        | 	local end_rel = pose_trans(pose_inv(p_center), scoop_end_pose)
        | 	local end_rel_tilted = pose_trans(end_rel, p[0, 0, 0, 0, ry, 0])
        | 	global tilted_pose_in_base = pose_trans(p_center, p[0,correction_y,correction_z,end_rel_tilted[3],end_rel_tilted[4], end_rel_tilted[5]])
        | 	global tilted_pose_in_base = pose_trans(tilted_pose_in_base, p[0, 0, spatula_len, 0, 0, 0])
        | 
        | 	if (Pow_name == "lactose_fine" or Pow_name == "Magnesium_sterate"):
        | 		tilt_send((angle_deg+5))
        | 	end
        | 	movel(tilted_pose_in_base, a=0.03, v=0.1)
        | 
        | 	if (Pow_name == "lactose_fine" or Pow_name == "Magnesium_sterate"):
        | 		tilt_send((angle_deg-5))
        | 	end
        | 
        | 	if (spatula=="spatula_flat_S" or spatula=="spatula_S"):
        | 		vibration_3()
        | 	else:
        | 		set_analog_out(0, vibration_voltage)
        | 	end
        | 	if (Pow_name=="Mannitol" or Pow_name =="NaCl"):
        | 		local n=1.4
        | 	else:
        | 		local n=1.5
        | 	end
        | 	local ry_level = deg2rad(ry_deg/n)
        | 	local end_rel_tilted_level = pose_trans(end_rel, p[0, 0, 0, 0, ry_level, 0])
        | 	local level_tilted_pose_in_base = pose_trans(p_center, p[0,correction_y,correction_z,end_rel_tilted_level[3],end_rel_tilted_level[4], end_rel_tilted_level[5]])
        | 	local level_tilted_pose_in_base = pose_trans(level_tilted_pose_in_base, p[0, 0, spatula_len, 0, 0, 0])
        | 
        | 	movel(level_tilted_pose_in_base, a=0.03, v=0.1)
        | 	#if (level>70.0):
        | 		#sleep(1.0)
        | 	#end
        | 	sleep(1.0)
        | 	#sleep(vibration_time)
        | 
        | 	movel(tilted_pose_in_base, a=0.03, v=0.1)
        | 	set_analog_out(0, 0.0)
        | 
        | 	tilt_pose_rel = pose_trans(pose_inv(p_center), tilted_pose_in_base)
        | 
        | 	lifted_pose_rel = pose_trans(lift_offset, tilt_pose_rel)
        | 
        | 	global lifted_pose = pose_trans(p_center, lifted_pose_rel)
        | 	movel(lifted_pose, a=0.03, v=0.1)
        | 	CCW_Rotate()
        | end
        | 
        | 
        | # calculate center pose on top of the container using pose transformation
        | def center_pose():
        | 	# pose transformation from side of the container to top to get center point
        | 	trans_rel = p[-0.005, 0.05, -0.027, 0, 0, 0]
        | 
        | 	p_translated = pose_trans(place_pose, trans_rel)
        | 	cx = p_translated[0]
        | 	cy = p_translated[1]
        | 	cz = p_translated[2]
        | 
        | 	global p_center_vertical = p[cx,cy,cz, 0, 0, 4.14]
        | 
        | 	#movej(p_center_vertical, a =0.3, v =0.3)
        | 	return p_center_vertical
        | end
        | 
        | # update center pose based on tilting
        | def updated_center_pose(p_center_vertical, angle_deg):
        | 	hinge_pose = pose_trans(p_center_vertical, p[0,0,-0.2,0,0,0])
        | 	local_rel = pose_trans(pose_inv(hinge_pose), p_center_vertical)
        | 
        | 	rot_tilt = p[0,0,0, -deg2rad(angle_deg),0,0]
        | 	local_rel_tilted = pose_trans(rot_tilt, local_rel)
        | 
        | 	global p_center = pose_trans(hinge_pose, local_rel_tilted)
        | 	return p_center
        | end
        | 
        | #------
        | # POTS commands
        | def tilt_send(angle):
        | 	socket_open("192.168.12.101", 80)
        | 	angle = 92.0 - angle
        | 	socket_send_string("Tilt,"+to_str(angle)+",0")
        | 	sync()
        | 	sleep(0.5)
        | 	socket_close()
        | end
        | 
        | def Motors_off():
        | 	socket_open("192.168.12.101", 80)
        | 	socket_send_string("Off,0,0")
        | 	sync()
        | 	sleep(0.5)
        | 	socket_close()
        | end
        | 
        | def Rotate():
        | 	socket_open("192.168.12.101", 80)
        | 	socket_send_string("FullRotation, 1, 2000")
        | 	sync()
        | 	sleep(0.5)
        | 	socket_close()
        | end
        | 
        | 
        | def CCW_Rotate():
        | 	socket_open("192.168.12.101", 80)
        | 	socket_send_string("FullRotation, -1, 2000")
        | 	sync()
        | 	sleep(0.5)
        | 	socket_close()
        | end
        | 
        | def tilt_to_home():
        | 	socket_open("192.168.12.101", 80)
        | 	socket_send_string("Home,0,0")
        | 	sync()
        | 	sleep(0.5)
        | 	socket_close()
        | end
    SuppressedNode
      Script file /programs/04 Scripts/dosing.script
        | def vibration_2():
        | 	set_analog_out(0,0.4)
        | 	sleep(0.8)
        | 	set_analog_out(0,0.0)
        | 	sleep(0.2)
        | end
        | 
        | def vibration_3():
        | 	set_analog_out(0,0.4)
        | 	sleep(0.5)
        | 	set_analog_out(0,0.0)
        | 	sleep(0.3)
        | end
        | 
        | def vibration_4():
        | 	set_analog_out(0,0.4)
        | 	sleep(0.6)
        | 	set_analog_out(0, 0.0)
        | 	sleep(0.5)
        | end
        | 
        | def vibration_1():
        | 	set_analog_out(0,0.4)
        | 	sleep(1)
        | 	set_analog_out(0,0.0)
        | 	sleep(0)
        | end
        | 
        | def move_tilt_in_steps(Pow_center, final_pose, steps):
        | 	i = 0
        | 	while i <= steps:
        | 		ratio = i / steps
        | 		pose_step = p[Pow_center[0] + ratio * (final_pose[0] - Pow_center[0]), Pow_center[1] + ratio * (final_pose[1] -Pow_center[1]),Pow_center[2] + ratio * (final_pose[2] - Pow_center[2]), Pow_center[3] + ratio * (final_pose[3] - Pow_center[3]), Pow_center[4] + ratio * (final_pose[4] - Pow_center[4]), Pow_center[5] + ratio * (final_pose[5] - Pow_center[5])]
        | 		movej(pose_step, a=1.2, v=0.15)
        | 		sleep(0.1)
        | 		i = i+1
        | 	end
        | end
        | 
        | def tilt_container(angle):
        | 	p_center = get_actual_tcp_pose()
        | 	hinge_offset = p[0,0,-0.23,0,0,0]
        | 	pivot_pose = pose_trans(p_center, hinge_offset)
        | 	pose_rel = pose_trans(pose_inv(pivot_pose), p_center)
        | 	angle_mid = (angle/2.0)*3.1416/180
        | 	angle_end = angle*3.1416/180
        | 	tilt_mid = p[0,0,0, -angle_mid, 0, 0]
        | 	tilt_end = p[0,0,0, -angle_end, 0, 0]
        | 	pose_rel_mid = pose_trans(tilt_mid, pose_rel)
        | 	pose_rel_end = pose_trans(tilt_end, pose_rel)
        | 	via_pose = pose_trans(pivot_pose, pose_rel_mid)
        | 	end_pose = pose_trans(pivot_pose, pose_rel_end)
        | 	movec(via_pose, end_pose, a=0.05, v=0.01, r=0.001)
        | 	p_center = get_actual_tcp_pose()
        | end
        | 
        | def deg2rad(d):
        | 	return d*3.141592/180
        | end
        | 
        | def map_tilt_to_ry_deg(container_deg):
        | 	#ry_deg = -0.875*container_deg +87.0
        | 	#return clamp(ry_deg, 5.0, 80.0)
        | 	if (Pow_name == "NaCl" or Pow_name == "Mannitol" or Pow_name == "CCS" or Pow_name == "MCC"):
        | 		if ( level>=10.0):
        | 			ry_min = 10.0
        | 			ry_max = 75.0
        | 		elif (level<10.00 and level >1.00):
        | 			ry_min = 16.0
        | 			ry_max = 65.0
        | 		else:
        | 			ry_min=17.0
        | 			ry_max=75.0
        | 		end
        | 	else:
        | 		if ( level>=10.0):
        | 			ry_min = 0.0
        | 			ry_max = 65.0
        | 		elif (level<10.00 and level >1.00):
        | 			ry_min = 10.0
        | 			ry_max = 45.0
        | 		else:
        | 			ry_min=0.0
        | 			ry_max=50.0
        | 		end
        | 
        | 	end
        | 	local span_count = angle_max -angle_min
        | 	local span_ry = ry_max - ry_min
        | 
        | 	local t = (container_deg -angle_min)/span_count
        | 	local ry_deg = ry_max - t*span_ry
        | 
        | 	return clamp(ry_deg, ry_min, ry_max)
        | 
        | end
        | 
        | def caluclate_corrections(level):
        | 	z_high = 0.01
        | 	z_low = -0.08
        | 	y_high = -0.01
        | 	y_low = -0.015
        | 
        | 	scale = (level - 10.0) / (100.0-10.0)
        | 
        | 	global correction_z = z_low + scale*(z_high - z_low)
        | 	global correction_y = y_low + scale*(y_high -y_low)
        | 
        | end
        | 
        | def scoop_powder(p_center):
        | 	#lift_offset = p[0, 0, 0.05, 0, 0, 0]
        | 	vibration_voltage = 0.4
        | 	vibration_time = 3.0
        | 	diameter = 0.07
        | 	global scoop_radius_default = 0.0
        | 	#p_center = center_pose_t
        | 
        | 
        | 	if (level >=70.00):
        | 		approach_offset = p[0.008,0,0.22,0,0,0]
        | 		lift_offset = p[0, 0, 0.05, 0, 0, 0]
        | 		caluclate_corrections(level)
        | 	elif (level >=10.00 and level <70):
        | 		approach_offset = p[0.008,0,0.22,0,0,0]
        | 		lift_offset = p[0, 0, 0.15, 0, 0, 0]
        | 		caluclate_corrections(level)
        | 	elif (level<10.00 and level >= 1.00):
        | 		approach_offset = p[0.01,0,0.22,0,0,0]
        | 		correction_z = -0.08
        | 		correction_y = -0.01
        | 		lift_offset = p[0, 0, 0.14, 0, 0, 0]
        | 	else:
        | 		approach_offset = p[0.008,0,0.22,0,0,0]
        | 		correction_z = -0.08
        | 		correction_y = -0.01
        | 		lift_offset = p[0, 0, 0.14, 0, 0, 0]
        |  	end
        | 
        | 	if (spatula == "spatula_L"):
        | 		global spatula_depth = 0.015
        | 	elif (spatula == "spatula_M"):
        | 		global spatula_depth = 0.01
        | 	elif (spatula == "spatula_S"):
        | 		global spatula_depth = 0.008
        | 	elif (spatula == "spatula_flat_M"):
        | 		global spatula_depth = 0.001
        | 	elif (spatula == "spatula_flat_S"):
        | 		global spatula_depth = 0.005
        | 	end
        | 
        | 	scoop_radius_default = diameter/2 - spatula_depth
        | 	scoop_entry_pose = pose_trans(p_center, approach_offset)
        | 	movel(scoop_entry_pose, a=0.1, v=0.25)
        | 
        | 	scoop_start_rel = p[scoop_radius_default, 0, scoop_depth, 0, 0, 0]
        | 
        | 	rot_mid = p[0, 0, 0, 0, 0, 0.785]
        | 	rot_end = p[0, 0, 0, 0, 0, 1.5708]
        | 
        | 	scoop_via_rel = pose_trans(rot_mid, scoop_start_rel)
        | 	scoop_end_rel = pose_trans(rot_end, scoop_start_rel)
        | 
        | 	scoop_start_pose = pose_trans(p_center, scoop_start_rel)
        | 	scoop_via_pose = pose_trans(p_center, scoop_via_rel)
        | 	scoop_end_pose = pose_trans(p_center, scoop_end_rel)
        | 
        | 	movel(scoop_start_pose, a=0.5, v=0.3)
        | 	#movel(p_center, a=0.5, v=1.0)
        | 	#sleep(5.0)
        | 
        | 	if (level<90.0):
        | 		Rotate()
        | 	end
        | 
        | 	#movec(scoop_via_pose, scoop_end_pose, a=0.03, v=0.05)
        | 	movec(scoop_via_pose, scoop_end_pose, a=0.03, v=0.02)
        | 	#movel(pose_trans(get_actual_tcp_pose(), p[0,0,0,0,0,deg2rad(90.0)]), a=0.03, v=0.05)
        | 	sleep(1.0)
        | 	local ry_deg = map_tilt_to_ry_deg(angle_deg)
        | 	local ry = deg2rad(ry_deg)
        | 	local end_rel = pose_trans(pose_inv(p_center), scoop_end_pose)
        | 	local end_rel_tilted = pose_trans(end_rel, p[0, 0, 0, 0, ry, 0])
        | 	global tilted_pose_in_base = pose_trans(p_center, p[0,correction_y,correction_z,end_rel_tilted[3],end_rel_tilted[4], end_rel_tilted[5]])
        | 	global tilted_pose_in_base = pose_trans(tilted_pose_in_base, p[0, 0, spatula_len, 0, 0, 0])
        | 
        | 	if (Pow_name == "lactose_fine" or Pow_name == "Magnesium_sterate"):
        | 		tilt_send((angle_deg+5))
        | 	end
        | 	movel(tilted_pose_in_base, a=0.03, v=0.1)
        | 
        | 	if (Pow_name == "lactose_fine" or Pow_name == "Magnesium_sterate"):
        | 		tilt_send((angle_deg-5))
        | 	end
        | 
        | 	if (spatula=="spatula_flat_S" or spatula=="spatula_S"):
        | 		vibration_3()
        | 	else:
        | 		set_analog_out(0, vibration_voltage)
        | 	end
        | 	if (Pow_name=="Mannitol" or Pow_name =="NaCl"):
        | 		local n=1.4
        | 	else:
        | 		local n=1.5
        | 	end
        | 	local ry_level = deg2rad(ry_deg/n)
        | 	local end_rel_tilted_level = pose_trans(end_rel, p[0, 0, 0, 0, ry_level, 0])
        | 	local level_tilted_pose_in_base = pose_trans(p_center, p[0,correction_y,correction_z,end_rel_tilted_level[3],end_rel_tilted_level[4], end_rel_tilted_level[5]])
        | 	local level_tilted_pose_in_base = pose_trans(level_tilted_pose_in_base, p[0, 0, spatula_len, 0, 0, 0])
        | 
        | 	movel(level_tilted_pose_in_base, a=0.03, v=0.1)
        | 	#if (level>70.0):
        | 		#sleep(1.0)
        | 	#end
        | 	sleep(1.0)
        | 	#sleep(vibration_time)
        | 
        | 	movel(tilted_pose_in_base, a=0.03, v=0.1)
        | 	set_analog_out(0, 0.0)
        | 
        | 	tilt_pose_rel = pose_trans(pose_inv(p_center), tilted_pose_in_base)
        | 
        | 	lifted_pose_rel = pose_trans(lift_offset, tilt_pose_rel)
        | 
        | 	global lifted_pose = pose_trans(p_center, lifted_pose_rel)
        | 	movel(lifted_pose, a=0.03, v=0.1)
        | 	CCW_Rotate()
        | end
        | 
        | 
        | def center_pose():
        | 	trans_rel = p[-0.005, 0.05, -0.015, 0, 0, 0]
        | 
        | 	p_translated = pose_trans(place_pose, trans_rel)
        | 	cx = p_translated[0]
        | 	cy = p_translated[1]
        | 	cz = p_translated[2]
        | 
        | 	global p_center_vertical = p[cx,cy,cz, 0, 0, 4.09]
        | 
        | 	#movej(p_center_vertical, a =0.3, v =0.3)
        | 	return p_center_vertical
        | end
        | 
        | def updated_center_pose(p_center_vertical, angle_deg):
        | 	hinge_pose = pose_trans(p_center_vertical, p[0,0,-0.2,0,0,0])
        | 	local_rel = pose_trans(pose_inv(hinge_pose), p_center_vertical)
        | 
        | 	rot_tilt = p[0,0,0, -deg2rad(angle_deg),0,0]
        | 	local_rel_tilted = pose_trans(rot_tilt, local_rel)
        | 
        | 	global p_center = pose_trans(hinge_pose, local_rel_tilted)
        | 	return p_center
        | end
        | 
        | def tilt_send(angle):
        | 	socket_open("192.168.12.101", 80)
        | 	angle = 92.0 - angle
        | 	socket_send_string("Tilt,"+to_str(angle)+",0")
        | 	sync()
        | 	sleep(0.5)
        | 	socket_close()
        | end
        | 
        | def Motors_off():
        | 	socket_open("192.168.12.101", 80)
        | 	socket_send_string("Off,0,0")
        | 	sync()
        | 	sleep(0.5)
        | 	socket_close()
        | end
        | 
        | def Rotate():
        | 	socket_open("192.168.12.101", 80)
        | 	socket_send_string("FullRotation, 1, 2000")
        | 	sync()
        | 	sleep(0.5)
        | 	socket_close()
        | end
        | 
        | 
        | def CCW_Rotate():
        | 	socket_open("192.168.12.101", 80)
        | 	socket_send_string("FullRotation, -1, 2000")
        | 	sync()
        | 	sleep(0.5)
        | 	socket_close()
        | end
        | def tilt_to_home():
        | 	socket_open("192.168.12.101", 80)
        | 	socket_send_string("Home,0,0")
        | 	sync()
        | 	sleep(0.5)
        | 	socket_close()
        | end
    Script file /programs/04 Scripts/Powder_all.script
      | global SERVER_IP   = "192.168.12.139"
      | global SERVER_PORT = 3002
      | 
      | global container_id = 0
      | global powder_id  = 0
      | global bulk_density = 0
      | global H          = 0
      | global H_c          = 0
      | global mouth_d     = 0
      | global mouth_sh    = 0
      | global length_c     = 0
      | global diameter   = 0
      | global empty_weight_g  = 0
      | global volume_ml    = 0
      | global shape_code   = 0
      | global flow_code   = 0
      | global shape = ""
      | global Flowability = ""
      | global full_weight_g = 0
      | global cent_edge = 0
      | global pick_2_base = 0.2 # distance from tcp to base of picking table
      | global wall_thickness = 0.001
      | 
      | def read_db_data():
      | 
      |   socket_open(SERVER_IP, SERVER_PORT)
      |   sleep(0.5)
      |   socket_send_string("GET_DATACODE_FLOATS")
      |   sleep(5)
      | 
      |   local fl = socket_read_ascii_float(14)
      |   socket_close()
      | 
      |   global container_id = fl[1]
      |   global powder_id = fl[2]
      |   global bulk_density = fl[3]
      |   global H          = fl[4]/1000
      |   global H_c          = fl[5]/1000
      |   global mouth_d     = fl[6]/1000
      |   global mouth_sh    = fl[7]/1000
      |   global length_c     = fl[8]/1000
      |   global diameter   = fl[9]/1000
      |   global empty_weight_g = fl[10]
      |   global volume_ml    = fl[11]
      |   global full_weight_g = fl[12]
      |   global flow_code   = fl[13]
      |   global shape_code   = fl[14]
      | 
      | 	if (flow_code == 1.0):
      | 	  global Flowability = "MEDIUM"
      | 	elif (flow_code == 2.0):
      | 	  global Flowability = "LOW"
      | 	else:
      | 	  global Flowability = "HIGH"
      | 	end
      | 
      |   if ( shape_code == 1.0):
      | 	shape = "cylindrical"
      | 	cent_edge =  diameter
      |   else:
      | 	shape = "cubical"
      | 	cent_edge =  length_c
      |   end
      | 
      | end
      | 
      | 
      | def send_picking_info(Pow_name, target_weight):
      |   socket_open(SERVER_IP, SERVER_PORT)
      |   cmd = "PICK:"+Pow_name+";"+to_str(target_weight)
      |   socket_send_string(cmd)
      |   sleep(0.1)
      |   socket_close()
      | end
      | 
      | #### POTS ####
      | def tilt_send(angle):
      | 	socket_open("192.168.12.101", 80)
      | 	angle = 90.0 - angle
      | 	socket_send_string("Tilt,"+to_str(angle)+",0")
      | 	sync()
      | 	sleep(0.5)
      | 	socket_close()
      | end
      | 
      | def Motors_off():
      | 	socket_open("192.168.12.101", 80)
      | 	socket_send_string("Off,0,0")
      | 	sync()
      | 	sleep(0.5)
      | 	socket_close()
      | end
      | 
      | def Rotate():
      | 	socket_open("192.168.12.101", 80)
      | 	socket_send_string("FullRotation, 1, 2000")
      | 	sync()
      | 	sleep(0.5)
      | 	socket_close()
      | end
      | 
      | def CCW_Rotate():
      | 	socket_open("192.168.12.101", 80)
      | 	socket_send_string("FullRotation, -1, 2000")
      | 	sync()
      | 	sleep(0.5)
      | 	socket_close()
      | end
      | 
      | def tilt_to_home():
      | 	socket_open("192.168.12.101", 80)
      | 	socket_send_string("Home,0,0")
      | 	sync()
      | 	sleep(0.5)
      | 	socket_close()
      | end
      | #######
      | def vibration_1():
      | 	set_analog_out(0,0.4)
      | 	sleep(1)
      | 	set_analog_out(0,0.0)
      | 	sleep(0)
      | end
      | 
      | def vibration_2():
      | 	set_analog_out(0,0.4)
      | 	sleep(0.8)
      | 	set_analog_out(0,0.0)
      | 	sleep(0.2)
      | end
      | 
      | def vibration_3():
      | 	set_analog_out(0,0.4)
      | 	sleep(0.5)
      | 	set_analog_out(0,0.0)
      | 	sleep(0.3)
      | end
      | 
      | def vibration_4():
      | 	set_analog_out(0,0.8)
      | 	sleep(0.6)
      | 	set_analog_out(0, 0.0)
      | 	sleep(0.5)
      | end
      | 
      | ##################
      | 
      | global gear_2_holder = 0.018
      | global gain_per_percent = 0.5
      | global w_dosed_total = 0.0
      | global last_scale = 0.0
      | global tilt_angle_sent = 0.0
      | global level = 0.0
      | global target_g = 0.0
      | global angle_max = 60
      | global angle_min = 10
      | global hinge_2_base = 0.0421
      | global TCP_2_tip_x = 0.0047
      | global spatula_len = 0.182
      | global spatula_offset = p[TCP_2_tip_x,0,spatula_len,0,0,0]
      | global SPATULA_L_VOL_ML = 5.0        # 1 teaspoon = 5 mL
      | global SPATULA_M_VOL_ML = 1.25       # 1/4 teaspoon = 1.25 mL
      | global SPATULA_S_VOL_ML = 0.15625    # 1/32 teaspoon = 0.15625 mL
      | global SPATULA_FLAT_M_VOL_ML  = 2.2
      | global SPATULA_FLAT_S_VOL_ML  = 1.2   #based on caluclations using rho = m/V
      | global ry_deg_safe = 0
      | global ry_deg = 0
      | 
      | 
      | 
      | def clamp(x, lo, hi):
      | 	if(x<lo):
      | 		return lo
      | 	elif (x>hi):
      | 		return hi
      | 	else:
      | 		return x
      | 	end
      | end
      | 
      | def compute_level_percent(W_now, weight_value):   # W_now = container+powder, weight_value = live scale reading
      |     local delta = weight_value - last_scale
      | 
      |     if (delta < 0.0):
      |         delta = 0.0
      |     end
      | 
      |     global w_dosed_total = w_dosed_total + delta
      |     global last_scale = weight_value     # update the last scale reading
      | 
      |     local W_eff = W_now - w_dosed_total
      |     if (W_eff <  empty_weight_g):
      |         W_eff =  empty_weight_g
      |     end
      | 
      |     # Compute powder level %
      |     level = 100.0 * (W_eff -  empty_weight_g) / (full_weight_g -  empty_weight_g)
      | 
      |     # Clamp to 0–100
      |     level = clamp(level, 0, 100)
      |   textmsg("deb 1 = ", level)
      |     return level
      | end
      | 
      | def deg2rad(d):
      | 	return d*3.141592/180
      | end
      | 
      | def my_abs(val):
      | 	if (val<0):
      | 		return -val
      | 	else:
      | 		return val
      | 	end
      | end
      | 
      | def compute_tilt_deg(level_percent):
      | 	angle = angle_min + gain_per_percent*(100.0-level_percent)
      | 
      |   	textmsg("deb 2 = ", angle)
      | 	return clamp(angle, angle_min, angle_max)
      | end
      | 
      | def tilt(level_percentage):
      | 	new_angle = compute_tilt_deg(level_percentage)
      | 	global angle_rel = new_angle - tilt_angle_sent
      | 
      | 	if my_abs(angle_rel)>2.0:
      | 		tilt_send(new_angle)
      | 		global angle_deg = new_angle
      | 		global tilt_angle_sent = new_angle
      | 		global p_center_vertical = center_pose()
      | 		global p_center = updated_center_pose(p_center_vertical, angle_deg)
      | 	end
      | 
      | 	if (level_percentage<85.0):
      | 		tilt_send(angle_deg)
      | 	end
      | end
      | 
      | def compute_scoop_depth(level):
      |   return ((100.0-level)/100.0)*(H -mouth_sh )
      | end
      | 
      | def map_tilt_to_ry_deg(container_deg, level):
      | 
      | 	if (Flowability == "HIGH" or Flowability == "MEDIUM"):
      | 		global scoop_depth = compute_scoop_depth(level)
      | 		safe_scoop_pivot = (mouth_d  - spatula_depth)/(scoop_depth+mouth_sh )
      | 		global ry_deg_safe = asin(safe_scoop_pivot)
      | 		global ry_deg = 90-container_deg
      | 	else:
      | 		global scoop_depth = compute_scoop_depth(level)
      | 		safe_scoop_pivot = (mouth_d  - spatula_depth)/(scoop_depth+mouth_sh )
      | 		global ry_deg_safe = asin(safe_scoop_pivot)
      | 		global ry_deg = 90-container_deg
      | 	end
      | 	return [ry_deg_safe,ry_deg]
      | end
      | 
      | def get_scoop_weight(spatula, bulk_density):
      | 
      | 	local vol = 0
      | 
      | 	if (spatula == "spatula_L"):
      | 		vol = SPATULA_L_VOL_ML
      | 		global spatula_depth = 0.015
      | 		global spatula_mid   = 0.016
      | 		global spatula_ry    = 0.0
      | 
      | 	elif (spatula == "spatula_M"):
      | 		vol = SPATULA_M_VOL_ML
      | 		global spatula_depth = 0.010
      | 		global spatula_mid   = 0.0105
      | 		global spatula_ry    = 0.0
      | 
      | 	elif (spatula == "spatula_S"):
      | 		vol = SPATULA_S_VOL_ML
      | 		global spatula_depth = 0.008
      | 		global spatula_mid   = 0.0063
      | 		global spatula_ry    = 0.0
      | 
      | 	elif (spatula == "spatula_flat_M"):
      | 		vol = SPATULA_FLAT_M_VOL_ML
      | 		global spatula_depth = 0.001
      | 		global spatula_mid   = 0.002
      | 		global spatula_ry    = 10.0
      | 
      | 	elif (spatula == "spatula_flat_S"):
      | 		vol = SPATULA_FLAT_S_VOL_ML
      | 		global spatula_depth = 0.005
      | 		global spatula_mid   = 0.016
      | 		global spatula_ry    = 2.0
      | 
      | 	else:
      | 		textmsg("Unknown spatula type")
      | 		return 0.0
      | 	end
      | 	global target_g = vol * bulk_density
      | 	return target_g
      | 
      | end
      | 
      | def select_spatula(Flowability, level, diff, bulk_density, mouth_d ):
      | 
      |     local k = 1.1
      | 
      |     global powder_height = (H  - mouth_sh ) * level/100
      | 
      |     # =====================================================
      |     # LOW FLOWABILITY
      |     # =====================================================
      |     if (Flowability == "LOW"):
      | 
      |         local gFM = get_scoop_weight("spatula_flat_M", bulk_density)
      | 
      |         local level_ok_FM = (spatula_mid * 2 < powder_height)
      |         local diff_ok_FM  = (diff > k * gFM)
      | 
      |         local flatM_ok = level_ok_FM and diff_ok_FM
      | 
      |         if (flatM_ok):
      |             return "spatula_flat_M"
      |         else:
      |             return "spatula_flat_S"
      |         end
      | 
      |     end
      | 
      | 
      |     # =====================================================
      |     # LARGE
      |     # =====================================================
      |     local gL = get_scoop_weight("spatula_L", bulk_density)
      | 
      |     local mouth_ok_L = (mouth_d  >= 0.05)
      |     local level_ok_L = (spatula_mid * 2 < powder_height)
      |     local diff_ok_L  = (diff > k * gL)
      | 
      |     local large_ok = mouth_ok_L and level_ok_L and diff_ok_L
      | 
      | 
      |     # =====================================================
      |     # MEDIUM
      |     # =====================================================
      |     local gM = get_scoop_weight("spatula_M", bulk_density)
      | 
      |     local level_ok_M = (spatula_mid * 2 < powder_height)
      |     local diff_ok_M  = (diff > k * gM)
      | 
      |     local medium_ok = level_ok_M and diff_ok_M
      | 
      | 
      |     # =====================================================
      |     # FINAL SELECTION
      |     # =====================================================
      |     if (large_ok):
      |         return "spatula_L"
      | 
      |     elif (medium_ok):
      |         return "spatula_M"
      | 
      |     else:
      |         return "spatula_S"
      |     end
      | 
      | end
      | 
      | def after_scoop():
      | 	tilt_send(angle_deg)
      | 	sleep(0.5)
      | 	movel(lifted_pose, a=0.05, v=0.2)
      | 	movel(tilted_pose_in_base2, a=0.05, v=0.2)
      | 	set_analog_out(0,0.4)
      | 	movel(pose_trans(tilted_pose_in_base2, p[0,0,0,0,0,2.0]), a=0.05, v=0.2)
      | 	set_analog_out(0,0.0)
      | 	movel(lifted_pose, a=0.05, v=0.2)
      | 	tilt_to_home()
      | end
      | 
      | def center_pose():
      | 	global p_translated = container_place
      | 	#global p_translated = pots_axis_temp
      | 
      | 	#cx = p_translated[0]
      | 	#cy = p_translated[1]
      | 	#cz = p_translated[2]
      | 
      | 	global p_center_vertical_temp = pose_trans(p_translated, p[0,0,0, deg2rad(90), 0, 0])
      | 	cx = p_center_vertical_temp[0]
      | 	cy = p_center_vertical_temp[1]
      | 	cz = p_center_vertical_temp[2]
      | 	#rx = p_center_vertical_temp[3]
      | 	#ry = p_center_vertical_temp[4]
      | 	rz = p_center_vertical_temp[5]
      | 
      | 	global p_center_vertical_temp = p[cx,cy,cz, 0, 0, rz]
      | 	trans_rel = p[0,0,-pick_2_base+H,0,0,0]
      | 	global p_center_vertical =  pose_trans(p_center_vertical_temp, trans_rel)
      | 	return p_center_vertical
      | end
      | 
      | def updated_center_pose(p_center_vertical, angle_deg):
      | 	hinge_pose = pose_trans(p_center_vertical, p[0,0,-hinge_2_base-gear_2_holder-H ,0,0,0])
      | 	local_rel = pose_trans(pose_inv(hinge_pose), p_center_vertical)
      | 
      | 	rot_tilt = p[0,0,0, -deg2rad(angle_deg),0,0]
      | 	local_rel_tilted = pose_trans(rot_tilt, local_rel)
      | 
      | 	global p_center = pose_trans(hinge_pose, local_rel_tilted)
      | 	return p_center
      | end
      | 
      | def scoop_powder(p_center):
      | 	vibration_voltage = 0.4
      | 	vibration_time = 3.0
      | 	global scoop_radius_default = 0.0
      | 
      | 
      | 	scoop_radius_default = mouth_d /2 - spatula_depth
      | 	scoop_safe_entry_pose = pose_trans(p_center, p[-TCP_2_tip_x,0,spatula_len+0.05,0,0,0])
      | 	scoop_entry_pose = pose_trans(p_center, p[-TCP_2_tip_x,0,spatula_len,0,0,0])
      | 
      | 	movel(scoop_safe_entry_pose, a=0.1, v=0.25)
      | 	movel(scoop_entry_pose, a=0.1, v=0.25)
      | 
      | 	scoop_start_rel_int = p[0, 0, -mouth_sh , 0, 0, 0]
      | 	scoop_start_pose_int = pose_trans(scoop_entry_pose, scoop_start_rel_int)
      | 
      | 	movel(scoop_start_pose_int, a=0.1, v=0.25)
      | 
      | 	if (spatula_mid * 2 < powder_height and spatula == "spatula_M" or spatula == "spatula_L"):
      | 
      | 		global total_depth = mouth_sh + scoop_depth + spatula_mid
      | 		global total_depth = clamp(total_depth, 0, H - spatula_mid)
      | 		scoop_start_rel = p[scoop_radius_default, 0, -total_depth, 0, 0, 0]
      | 
      | 		rot_mid = p[0, 0, 0, 0, 0, 0.785]
      | 		rot_end = p[0, 0, 0, 0, 0, 1.5708]
      | 
      | 		scoop_via_rel = pose_trans(rot_mid, scoop_start_rel)
      | 		scoop_end_rel = pose_trans(rot_end, scoop_start_rel)
      | 
      | 		scoop_start_pose = pose_trans(scoop_entry_pose, scoop_start_rel)
      | 		scoop_via_pose = pose_trans(scoop_entry_pose, scoop_via_rel)
      | 		scoop_end_pose = pose_trans(scoop_entry_pose, scoop_end_rel)
      | 
      | 		movel(scoop_start_pose, a=0.5, v=0.3)
      | 
      | 		if (level<90.0):
      | 			Rotate()
      | 		end
      | 
      | 		movec(scoop_via_pose, scoop_end_pose, a=0.03, v=0.02)
      | 		sleep(1.0)
      | 		#local ry_deg = map_tilt_to_ry_deg(angle_deg,level)
      | 		local ry_result = map_tilt_to_ry_deg(angle_deg,level)
      | 		global ry_safe = ry_result[0]
      | 		global ry = deg2rad(ry_result[1])
      | 
      | 		# safe_retention
      | 		local pivot_pose = pose_trans(scoop_end_pose, p[0,0,total_depth-spatula_len,0,0,0])
      | 		local end_rel = pose_trans(pose_inv(pivot_pose), scoop_end_pose)
      | 		local end_rel_tilted = pose_trans(end_rel, p[0, 0, 0, 0, ry_safe, 0])
      | 		global tilted_pose_in_base = pose_trans(pivot_pose, p[0,0,0,end_rel_tilted[3],end_rel_tilted[4], end_rel_tilted[5]])
      | 		global tilted_pose_in_base = pose_trans(tilted_pose_in_base, p[0, 0, spatula_len-total_depth, 0, 0, 0])
      | 		# sptula pivoted around the container rim of the mouth at ry_safe
      | 		movel(tilted_pose_in_base, a=0.03, v=0.1)
      | 
      | 		#popup("is the spatula crashing at front? ", blocking = True)
      | 		# safe_retention_above
      | 		# calculate x , z movements
      | 
      | 		global safe_x = sin(ry_safe)*(scoop_depth - (mouth_d -spatula_depth)/tan(90-ry_safe/2))
      | 		global safe_z = cos(ry_safe)*(scoop_depth - (mouth_d -spatula_depth)/tan(90-ry_safe/2))
      | 
      | 		local safe_up = pose_trans(tilted_pose_in_base, p[-safe_x,0,safe_z,0,0,0])
      | 		movel(safe_up, a=0.03, v=0.1)
      | 
      | 		#popup("is the spatula crashing at neck? ", blocking = True)
      | 
      | 		# full exit step by step
      | 		#local alpha = atan(2*mouth_sh /mouth_d )
      | 
      | 		#global cent_pose_cont_x = sin(ry_safe)*(scoop_depth - (mouth_d -spatula_depth)/tan(90-ry_safe/2))
      | 		#global cent_pose_cont_z = cos(ry_safe)*(scoop_depth+mouth_sh  - (mouth_d -spatula_depth)/tan(90-ry_safe/2))
      | 		#local cent_pose_cont = pose_trans(safe_up, p[])
      | 
      | 		# full exit
      | 		local pivot_pose2 = pose_trans(tilted_pose_in_base, p[0,0,total_depth-spatula_len,0,0,0])
      | 		local end_rel2 = pose_trans(pose_inv(pivot_pose2), tilted_pose_in_base)
      | 		#popup("is the spatula crashing front? ", blocking = True)
      | 		local end_rel_tilted2 = pose_trans(end_rel2, p[0, 0, 0, 0, ry-ry_safe, 0])
      | 		global tilted_pose_in_base2 = pose_trans(pivot_pose2, p[0,0,0,end_rel_tilted2[3],end_rel_tilted2[4], end_rel_tilted2[5]])
      | 		global tilted_pose_in_base2 = pose_trans(tilted_pose_in_base2, p[-TCP_2_tip_x, 0, spatula_len-scoop_radius_default-spatula_mid, 0, 0, 0])
      | 		# spaula exited at center of the mouth at ry
      | 		movel(tilted_pose_in_base2, a=0.03, v=0.1)
      | 		#popup("is the spatula crashing at mouth? ", blocking = True)
      | 
      | 	else : # emptying logic
      | 		spatula_base = pose_trans(scoop_entry_pose, p[0, 0, -H, 0, 0, 0])
      | 		local pivot_pose = pose_trans(scoop_entry_pose, p[0,0,-spatula_len,0,0,0])
      | 		# tilt inwards
      | 		global in_angle = atan((cent_edge-spatula_depth)/(2*H))
      | 		spatula_tilt_rel = pose_trans(pose_inv(pivot_pose), spatula_base)
      | 
      | 		spatula_tilt = pose_trans(spatula_tilt_rel, p[0, 0, 0, in_angle, 0, 0])
      | 		global tilted_pose = pose_trans(pivot_pose, p[0,0,0,spatula_tilt[3],spatula_tilt[4], spatula_tilt[5]])
      | 
      | 		global tilted_pose = pose_trans(tilted_pose, p[0,0,spatula_len-H,0,0,0])
      | 
      | 		movel(tilted_pose,a=0.1, v=0.25)
      | 		Rotate()
      | 
      | 		rot_mid = p[0, 0, 0, 0, 0, 0.785]
      | 		rot_end = p[0, 0, 0, 0, 0, 1.5708]
      | 
      | 		scoop_via_rel = pose_trans(tilted_pose, rot_mid)
      | 		scoop_end_rel = pose_trans(tilted_pose, rot_end)
      | 
      | 		movec(scoop_via_rel, scoop_end_rel, a=0.03, v=0.02)
      | 		popup("is the spatula crashing front? ", blocking = True)
      | 
      | 		scoop_via_pose = pose_trans(pivot_pose, scoop_via_rel)
      | 		scoop_end_pose = pose_trans(pivot_pose, scoop_end_rel)
      | 
      | 		#movec(scoop_via_pose, scoop_end_pose, a=0.03, v=0.02)
      | 		popup("is the spatula crashing front? ", blocking = True)
      | 		local ry_result = map_tilt_to_ry_deg(angle_deg,level)
      | 		global ry_safe = ry_result[0]
      | 		global ry = deg2rad(ry_result[1])
      | 
      | 		# full exit
      | 		#local pivot_pose2 = pose_trans(scoop_entry_pose, p[0,0,-spatula_len,0,0,0])
      | 		local end_rel2 = pose_trans(pose_inv(pivot_pose), scoop_end_pose)
      | 		popup("is the spatula crashing front? ", blocking = True)
      | 		local end_rel_tilted2 = pose_trans(end_rel2, p[0, 0, 0, 0, ry, 0])
      | 		global tilted_pose_in_base2 = pose_trans(pivot_pose, p[0,0,0,end_rel_tilted2[3],end_rel_tilted2[4], end_rel_tilted2[5]])
      | 		global tilted_pose_in_base2 = pose_trans(tilted_pose_in_base2, p[0, 0, spatula_len, 0, 0, 0])
      | 		# sptula exited at center of the mouth at ry
      | 		movel(tilted_pose_in_base2, a=0.03, v=0.1)
      | 		popup("is the spatula crashing at mouth? ", blocking = True)
      | 	end
      | 
      | 	if (spatula=="spatula_flat_S" or spatula=="spatula_S"):
      | 		vibration_3()
      | 	elif (spatula == "spatula_M"):
      | 		vibration_4()
      | 	else:
      | 		set_analog_out(0, vibration_voltage)
      | 	end
      | 
      | 	# remove excess
      | 	local pivot_pose_level = pose_trans(tilted_pose_in_base2, p[0,0,-spatula_len,0,0,0])
      | 	local end_rel_level = pose_trans(pose_inv(pivot_pose_level), tilted_pose_in_base2)
      | 	#local ry_level = ry/1.5
      | 	local ry_level = deg2rad(15)
      | 	local end_rel_tilted_level = pose_trans(end_rel_level, p[0, 0, 0, 0, -ry_level, 0])
      | 	local end_rel_tilted_level2 = pose_trans(pivot_pose_level, p[0, 0, 0,end_rel_tilted_level[3],end_rel_tilted_level[4], end_rel_tilted_level[5]])
      | 	local end_rel_tilted_level2 = pose_trans(end_rel_tilted_level2, p[0,0,spatula_len,0,0,0])
      | 	movel(end_rel_tilted_level2, a=0.03, v=0.1)
      | 
      | 	movel(tilted_pose_in_base2, a=0.03, v=0.1)
      | 	set_analog_out(0, 0.0)
      | 	#popup("safe out + moving towards beaker", title = "Pause", blocking = True)
      | 	global lifted_pose = pose_trans(tilted_pose_in_base2, p[-0.04,0,0.04,0,0,0]) # safety distance away from the container
      | 
      | 	movel(lifted_pose, a=0.03, v=0.1)
      | 	CCW_Rotate()
      | end
      | 
      | def auto_tilt_and_scoop(W_now, target_weight, weight_value):
      | 	global level = compute_level_percent(W_now, weight_value)
      | 
      | 	global spatula = select_spatula(Flowability, level, diff, bulk_density, mouth_d )
      | 	textmsg("deb 4 8 = ", spatula)
      | 	#global target_g = get_scoop_weight(spatula, bulk_density)
      | 
      |   	#textmsg("deb 4 = ", target_g)
      | 	#send_scoop_target_info()
      | 
      | 	global scoop_depth = compute_scoop_depth(level)
      | 
      |   	textmsg("deb 5 = ", scoop_depth)
      | 	tilt_to_home()
      | 	sleep(0.5)
      | 	tilt(level)
      | 	sleep(1.5)
      |   	#popup("is the pots tilted? ", blocking = True)
      |   	#textmsg("deb 6 = ", p_center)
      | 	scoop_powder(p_center)
      | 
      |   	textmsg("deb 7 - sucess")
      | end
    Script file /programs/04 Scripts/Weight_scale_socket_s.script
      | global s_depth = 0
      | global s_length =0
      | global s_volume = 0
      | global ry_theta  = 0
      | 
      | def get_weight():
      | 	socket_open(SERVER_IP,SERVER_PORT)
      | 	sleep(0.2)
      | 	textmsg("socket opened successfully!")
      | 	socket_send_string("GET_WEIGHT")
      | 	sleep(0.2)
      | 	sync()
      | 	sleep(0.2)
      | 	receiveFromServ = socket_read_ascii_float(6)
      | 	sleep(1)
      | 	#while (receiveFromServ[0] <1):
      | 		#receiveFromServ = socket_read_ascii_float(1)
      | 		#sleep(1)
      | 		#textmsg("retrying read:", receiveFromServ)
      | 	#end
      | 	textmsg("Received weight:", receiveFromServ[1])
      | 	sleep(0.2)
      | 	socket_close()
      | 	sleep(0.2)
      | 	return receiveFromServ[1]
      | end
      | 
      | def tare_scale():
      | 	socket_open(SERVER_IP,SERVER_PORT)
      | 	socket_send_string("TARE")
      | 	sleep(2)
      | 	socket_close()
      | end
      | 
      | def zero_scale():
      | 	socket_open(SERVER_IP,SERVER_PORT)
      | 	socket_send_string("ZERO")
      | 	sleep(0.5)
      | 	socket_close()
      | end
      | 
      | def log_weight():
      | 	socket_open(SERVER_IP,SERVER_PORT)
      | 	socket_send_string("LOG_WEIGHT")
      | 	sleep(0.5)
      | 	socket_close()
      | end
      | 
      | def send_target_info():
      | 	socket_open(SERVER_IP,SERVER_PORT)
      | 	socket_send_string("SET_TARGET:" + to_str(target_weight))
      | 	sleep(0.2)
      | 	socket_close()
      | end
      | def send_powder_info():
      | 	socket_open(SERVER_IP,SERVER_PORT)
      | 	socket_send_string("SET_POWDER:" + Pow_name)
      | 	sleep(0.2)
      | 	socket_close()
      | end
      | def send_spatula_info():
      | 	socket_open(SERVER_IP,SERVER_PORT)
      | 	socket_send_string("SET_SPATULA:" + spatula)
      | 	#sleep(1)
      | 
      | 	#local fl = socket_read_ascii_float(4)
      |   	#socket_close()
      | 
      |   	#global s_depth = fl[1]
      |   	#global s_length = fl[2]
      |  	#global s_volume = fl[3]
      |  	#global ry_theta  = fl[4]
      | 	sleep(0.2)
      | 
      | end
      | 
      | def send_level_info():
      | 	socket_open(SERVER_IP,SERVER_PORT)
      | 	socket_send_string("SET_LEVEL:" + to_str(level))
      | 	sleep(0.2)
      | 	socket_close()
      | end
      | def send_weight_info():
      |   socket_open(SERVER_IP, SERVER_PORT)
      |   #rq_open_and_wait()
      |   cmd = "GET_CONT_WEIGHT"
      |   socket_send_string(cmd)
      |   sync()
      |   sleep(0.5)
      |   receiveFromSer = socket_read_ascii_float(1)
      |   socket_close()
      |   return receiveFromSer[1]
      | end
  Folder BeforeStarts [hidden by the author, left out]
  Folder powder dispensing variable init [hidden by the author, left out]
Robot Program (runOnlyOnce=false)
  Folder MAIN [hidden by the author, left out]
Thread Thread_1 (runOnlyOnce=false)
  If Start_thread≟ True
    weight_value := get_weight()
    Wait Sleep waitTime=0.2
    Script: sync()
  Script: sync()
Thread Thread_2 (runOnlyOnce=false)
  Loop While (checkContinuously=true) expression=vib_thread≟ True
    diff := target_weight-weight_value
    If diff>0.02 and spatula≠"spatula_flat_S" (checkContinuously=true)
      SuppressedNode
        Script: vibration_1()
      Set AnalogOutput pin=analog_out[0]; analogValue=4
    ElseIf diff>0.02 and spatula≟"spatula_flat_S"
      Script: vibration_3()
    ElseIf diff≤0.03 (checkContinuously=true)
      Script: vibration_2()
    SuppressedNode
      ElseIf diff≥0.01 and diff<0.05
        Script: vibration_3()
    SuppressedNode
      ElseIf diff>0 and diff<0.01
        Script: vibration_4()
    Else 
      Set AnalogOutput pin=analog_out[0]; analogValue=0
  Script: sync()
SubProgram  [hidden by the author, left out]
SubProgram  [hidden by the author, left out]
SubProgram -> Sub_Action_V4
